{attribute 'no_assign'}
FUNCTION_BLOCK FB_LN_WTURBINE_LD0_WCNV1 EXTENDS FB_AcsiCommonLogicalNodeClass
VAR_INPUT
	Beh: FB_DO_WTURBINE_LD0_WCNV1_Beh := (sClass:='ENS', bLinkResult:=THIS^.AddDataToContainer(ipData:=Beh));
	Torq: FB_DO_WTURBINE_LD0_WCNV1_Torq := (sClass:='MV', bLinkResult:=THIS^.AddDataToContainer(ipData:=Torq));
END_VAR
VAR
END_VAR

END_FUNCTION_BLOCK

(* stored: Version 1.1.0.1
   POU FB_LN_WTURBINE_LD0_WCNV1: Id {8491b4d6-8485-4f48-8169-3efc00dc07ab}, SpecialFunc None *)
